FUNCTION_BLOCK FB_CIP_Source EXTENDS FB_SFC_Cycle IMPLEMENTS ITF_FB_SFC_Cycle
VAR_INPUT
	//eElementID			: E_Element_List;
	
	valTank_Water			: E_Pis_Name;
	valTank_R_Water			: E_Pis_Name;
	valTank_Detergent		: E_Pis_Name;
	valTank_DisInfection	: E_Pis_Name;	
	valDrain				: E_Pis_Name;
END_VAR
VAR_OUTPUT
END_VAR
VAR
	//refElement		: REFERENCE TO FB_Element;
	//refState_Long		: REFERENCE TO E_Element_State_Long;
	eReq				: E_CIP_Source;
	eProcess			: E_CIP_Source;
	eStatus				: E_CIP_Source;
	
	fbPis					: FB_Piston;
	stPis_Tank_Water		: REFERENCE TO ST_Piston;
	stPis_Tank_R_Water		: REFERENCE TO ST_Piston;
	stPis_Tank_Detergent	: REFERENCE TO ST_Piston;
	stPis_Tank_DisInfection	: REFERENCE TO ST_Piston;
	stPis_Drain				: REFERENCE TO ST_Piston;
	rt_Req_Reset: R_TRIG;
END_VAR
VAR_IN_OUT


END_VAR

act_GetReference();

act_Oper();
IF NOT Init.x THEN;
	act_Status();
END_IF

m_Request_Reset(memo:=rt_Req_Reset);//

ACTION _aClose_active:
bStepDone:=FALSE;
IF TRUE 
AND eStatus=E_CIP_Source.eClose
THEN;
	bStepDone:=TRUE;
END_IF
END_ACTION

ACTION _aClose_entry:
fbPis.m_SetByRecipe(stPis:=stPis_Tank_Water, 			req:=E_Piston_Recipe_State.Release);
fbPis.m_SetByRecipe(stPis:=stPis_Tank_R_Water, 			req:=E_Piston_Recipe_State.Release);
fbPis.m_SetByRecipe(stPis:=stPis_Tank_Detergent, 		req:=E_Piston_Recipe_State.Release);
fbPis.m_SetByRecipe(stPis:=stPis_Tank_DisInfection, 	req:=E_Piston_Recipe_State.Release);
fbPis.m_SetByRecipe(stPis:=stPis_Drain, 				req:=E_Piston_Recipe_State.Release);
END_ACTION

ACTION _aDetergent_entry:
fbPis.m_SetByRecipe(stPis:=stPis_Tank_Water, 			req:=E_Piston_Recipe_State.Release);
fbPis.m_SetByRecipe(stPis:=stPis_Tank_R_Water, 			req:=E_Piston_Recipe_State.Release);
fbPis.m_SetByRecipe(stPis:=stPis_Tank_Detergent, 		req:=E_Piston_Recipe_State.Act);
fbPis.m_SetByRecipe(stPis:=stPis_Tank_DisInfection, 	req:=E_Piston_Recipe_State.Release);
//fbPis.m_SetByRecipe(stPis:=stPis_Drain, 				req:=E_Piston_Recipe_State.Act);
END_ACTION

ACTION _aDone_entry:
eProcess:=E_CIP_Source.eNone;
eReq:=E_CIP_Source.eNone;
bRun:=FALSE;
bDone:=TRUE;
END_ACTION

ACTION _aInit_active:
SFCReset:=FALSE;
END_ACTION

ACTION _aInit_exit:
eProcess:=E_CIP_Source.eNone;
eReq:=E_CIP_Source.eNone;
END_ACTION

ACTION _aR_Water_entry:
fbPis.m_SetByRecipe(stPis:=stPis_Tank_Water, 			req:=E_Piston_Recipe_State.Release);
fbPis.m_SetByRecipe(stPis:=stPis_Tank_R_Water, 			req:=E_Piston_Recipe_State.Act);
fbPis.m_SetByRecipe(stPis:=stPis_Tank_Detergent, 		req:=E_Piston_Recipe_State.Release);
fbPis.m_SetByRecipe(stPis:=stPis_Tank_DisInfection, 	req:=E_Piston_Recipe_State.Release);
//fbPis.m_SetByRecipe(stPis:=stPis_Drain, 				req:=E_Piston_Recipe_State.Act);
END_ACTION

ACTION _aReady_active:


CASE eReq OF
	E_CIP_Source.eClose:;
			IF TRUE THEN;
				eProcess:=E_CIP_Source.eClose;
			END_IF

	E_CIP_Source.eT91_Sanitation:;
			IF TRUE THEN;
				eProcess:=E_CIP_Source.eT91_Sanitation;
			END_IF	
			
	E_CIP_Source.eT92_Detergent:;
			IF TRUE THEN;
				eProcess:=E_CIP_Source.eT92_Detergent;
			END_IF	

	E_CIP_Source.eT93_R_Water:;
			IF TRUE THEN;
				eProcess:=E_CIP_Source.eT93_R_Water;
			END_IF	
			
	E_CIP_Source.eT94_Water:;
			IF TRUE THEN;
				eProcess:=E_CIP_Source.eT94_Water;
			END_IF	

END_CASE
END_ACTION

ACTION _aReady_entry:

END_ACTION

ACTION _aReady_exit:
bRun:=TRUE;
bDone:=FALSE;
END_ACTION

ACTION _aSanitation_entry:
fbPis.m_SetByRecipe(stPis:=stPis_Tank_Water, 			req:=E_Piston_Recipe_State.Release);
fbPis.m_SetByRecipe(stPis:=stPis_Tank_R_Water, 			req:=E_Piston_Recipe_State.Release);
fbPis.m_SetByRecipe(stPis:=stPis_Tank_Detergent, 		req:=E_Piston_Recipe_State.Release);
fbPis.m_SetByRecipe(stPis:=stPis_Tank_DisInfection, 	req:=E_Piston_Recipe_State.Act);
END_ACTION

ACTION _aT91_Drain_Done_active:
bStepDone:=FALSE;
IF TRUE 
AND eStatus=E_CIP_Source.eT91_Sanitation
THEN;
	bStepDone:=TRUE;
END_IF
END_ACTION

ACTION _aT91_Drain_Done_entry:
fbPis.m_SetByRecipe(stPis:=stPis_Drain, 				req:=E_Piston_Recipe_State.Act);
END_ACTION

ACTION _aT92_Drain_Done_active:
bStepDone:=FALSE;
IF TRUE 
AND eStatus=E_CIP_Source.eT92_Detergent
THEN;
	bStepDone:=TRUE;
END_IF
END_ACTION

ACTION _aT92_Drain_Done_entry:
fbPis.m_SetByRecipe(stPis:=stPis_Drain, 				req:=E_Piston_Recipe_State.Act);
END_ACTION

ACTION _aT93_Drain_Done_active:
bStepDone:=FALSE;
IF TRUE 
AND eStatus=E_CIP_Source.eT93_R_Water
THEN;
	bStepDone:=TRUE;
END_IF
END_ACTION

ACTION _aT93_Drain_Done_entry:
fbPis.m_SetByRecipe(stPis:=stPis_Drain, 				req:=E_Piston_Recipe_State.Act);
END_ACTION

ACTION _aWater_active:
bStepDone:=FALSE;
IF TRUE 
AND eStatus=E_CIP_Source.eT94_Water
THEN;
	bStepDone:=TRUE;
END_IF
END_ACTION

ACTION _aWater_entry:
fbPis.m_SetByRecipe(stPis:=stPis_Tank_Water, 			req:=E_Piston_Recipe_State.Act);
fbPis.m_SetByRecipe(stPis:=stPis_Tank_R_Water, 			req:=E_Piston_Recipe_State.Release);
fbPis.m_SetByRecipe(stPis:=stPis_Tank_Detergent, 		req:=E_Piston_Recipe_State.Release);
fbPis.m_SetByRecipe(stPis:=stPis_Tank_DisInfection, 	req:=E_Piston_Recipe_State.Release);
fbPis.m_SetByRecipe(stPis:=stPis_Drain, 				req:=E_Piston_Recipe_State.Release);
END_ACTION

ACTION act_GetReference:
m_Set_SFCFlags_Reference();
//refElement REF= fbElement[eElementID];
//refState_Long REF= fbElement[eElementID].eState_Long;
	
stPis_Tank_Water			REF= g_Piston.stPis[valTank_Water];
stPis_Tank_R_Water			REF= g_Piston.stPis[valTank_R_Water];
stPis_Tank_Detergent		REF= g_Piston.stPis[valTank_Detergent];
stPis_Tank_DisInfection		REF= g_Piston.stPis[valTank_DisInfection];
stPis_Drain					REF= g_Piston.stPis[valDrain];
END_ACTION

ACTION act_Oper:
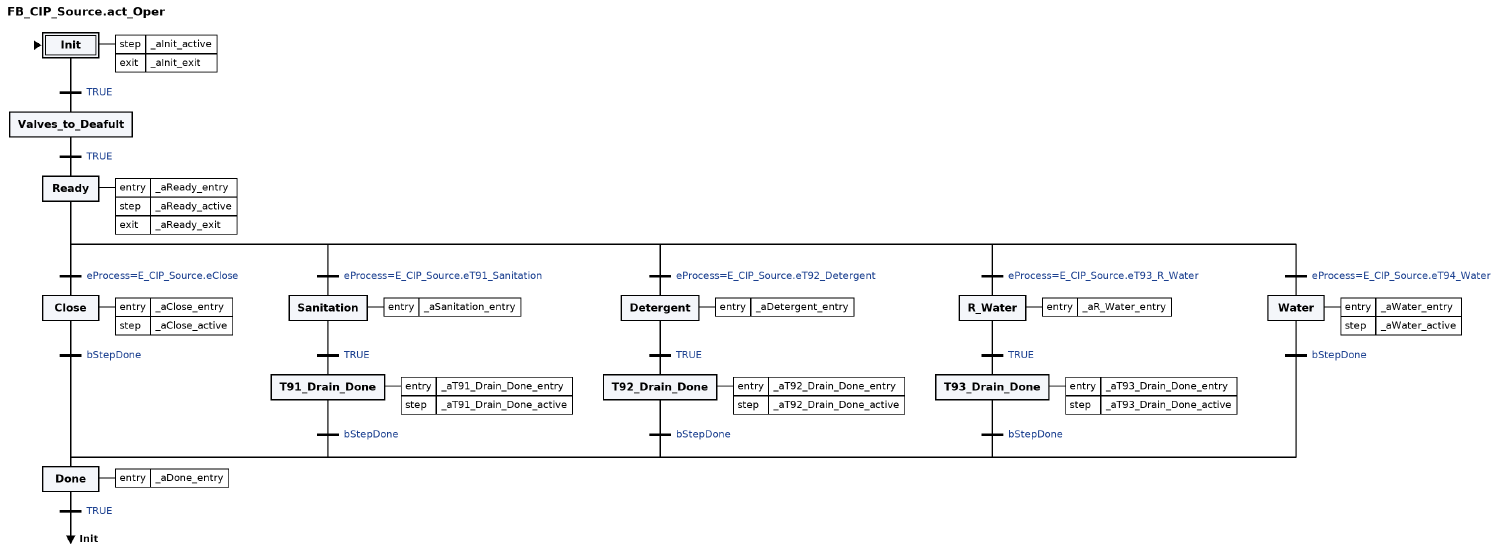
INITIAL_STEP Init:  // min time T#0.5s
    _aInit_active(N);  // step action
    _aInit_exit(P0);  // exit action
END_STEP
TRANSITION FROM Init TO Valves_to_Deafult
    := TRUE;
END_TRANSITION
STEP Valves_to_Deafult:
END_STEP
TRANSITION FROM Valves_to_Deafult TO Ready
    := TRUE;
END_TRANSITION
STEP Ready:
    _aReady_entry(P1);  // entry action
    _aReady_active(N);  // step action
    _aReady_exit(P0);  // exit action
END_STEP
TRANSITION FROM Ready TO Close
    := eProcess=E_CIP_Source.eClose;
END_TRANSITION
STEP Close:
    _aClose_entry(P1);  // entry action
    _aClose_active(N);  // step action
END_STEP
TRANSITION FROM Close TO Done
    := bStepDone;
END_TRANSITION
TRANSITION FROM Ready TO Sanitation
    := eProcess=E_CIP_Source.eT91_Sanitation;
END_TRANSITION
STEP Sanitation:  // min time T#7s
    _aSanitation_entry(P1);  // entry action
END_STEP
TRANSITION FROM Sanitation TO T91_Drain_Done
    := TRUE;
END_TRANSITION
STEP T91_Drain_Done:
    _aT91_Drain_Done_entry(P1);  // entry action
    _aT91_Drain_Done_active(N);  // step action
END_STEP
TRANSITION FROM T91_Drain_Done TO Done
    := bStepDone;
END_TRANSITION
TRANSITION FROM Ready TO Detergent
    := eProcess=E_CIP_Source.eT92_Detergent;
END_TRANSITION
STEP Detergent:  // min time T#6s
    _aDetergent_entry(P1);  // entry action
END_STEP
TRANSITION FROM Detergent TO T92_Drain_Done
    := TRUE;
END_TRANSITION
STEP T92_Drain_Done:
    _aT92_Drain_Done_entry(P1);  // entry action
    _aT92_Drain_Done_active(N);  // step action
END_STEP
TRANSITION FROM T92_Drain_Done TO Done
    := bStepDone;
END_TRANSITION
TRANSITION FROM Ready TO R_Water
    := eProcess=E_CIP_Source.eT93_R_Water;
END_TRANSITION
STEP R_Water:  // min time T#5s
    _aR_Water_entry(P1);  // entry action
END_STEP
TRANSITION FROM R_Water TO T93_Drain_Done
    := TRUE;
END_TRANSITION
STEP T93_Drain_Done:
    _aT93_Drain_Done_entry(P1);  // entry action
    _aT93_Drain_Done_active(N);  // step action
END_STEP
TRANSITION FROM T93_Drain_Done TO Done
    := bStepDone;
END_TRANSITION
TRANSITION FROM Ready TO Water
    := eProcess=E_CIP_Source.eT94_Water;
END_TRANSITION
STEP Water:
    _aWater_entry(P1);  // entry action
    _aWater_active(N);  // step action
END_STEP
TRANSITION FROM Water TO Done
    := bStepDone;
END_TRANSITION
STEP Done:  // min time T#0.2s
    _aDone_entry(P1);  // entry action
END_STEP
TRANSITION FROM Done TO Init
    := TRUE;
END_TRANSITION
// branch label Branch1_act_Oper
END_ACTION

ACTION act_Status:
IF bReady AND bDone OR TRUE THEN;
	IF TRUE 
	AND fbPis.m_CheckByRecipe(stPis:=stPis_Tank_Water, 			req:=E_Piston_Recipe_State.Release)
	AND fbPis.m_CheckByRecipe(stPis:=stPis_Tank_R_Water, 		req:=E_Piston_Recipe_State.Release)
	AND fbPis.m_CheckByRecipe(stPis:=stPis_Tank_Detergent, 		req:=E_Piston_Recipe_State.Release)
	AND fbPis.m_CheckByRecipe(stPis:=stPis_Tank_DisInfection, 	req:=E_Piston_Recipe_State.Release)
	AND fbPis.m_CheckByRecipe(stPis:=stPis_Drain, 				req:=E_Piston_Recipe_State.Release)
	THEN;
		eStatus:=E_CIP_Source.eClose;
	
	ELSIF TRUE 
	AND fbPis.m_CheckByRecipe(stPis:=stPis_Tank_Water, 			req:=E_Piston_Recipe_State.Act)
	AND fbPis.m_CheckByRecipe(stPis:=stPis_Tank_R_Water, 		req:=E_Piston_Recipe_State.Release)
	AND fbPis.m_CheckByRecipe(stPis:=stPis_Tank_Detergent, 		req:=E_Piston_Recipe_State.Release)
	AND fbPis.m_CheckByRecipe(stPis:=stPis_Tank_DisInfection, 	req:=E_Piston_Recipe_State.Release)
	AND fbPis.m_CheckByRecipe(stPis:=stPis_Drain, 				req:=E_Piston_Recipe_State.Release)
	THEN;
		eStatus:=E_CIP_Source.eT94_Water;
		
	ELSIF TRUE 
	AND fbPis.m_CheckByRecipe(stPis:=stPis_Tank_Water, 			req:=E_Piston_Recipe_State.Release)
	AND fbPis.m_CheckByRecipe(stPis:=stPis_Tank_R_Water, 		req:=E_Piston_Recipe_State.Act)
	AND fbPis.m_CheckByRecipe(stPis:=stPis_Tank_Detergent, 		req:=E_Piston_Recipe_State.Release)
	AND fbPis.m_CheckByRecipe(stPis:=stPis_Tank_DisInfection, 	req:=E_Piston_Recipe_State.Release)
	AND fbPis.m_CheckByRecipe(stPis:=stPis_Drain, 				req:=E_Piston_Recipe_State.Act)
	THEN;
		eStatus:=E_CIP_Source.eT93_R_Water;
		
	ELSIF TRUE 	
	AND fbPis.m_CheckByRecipe(stPis:=stPis_Tank_Water, 			req:=E_Piston_Recipe_State.Release)
	AND fbPis.m_CheckByRecipe(stPis:=stPis_Tank_R_Water, 		req:=E_Piston_Recipe_State.Release)
	AND fbPis.m_CheckByRecipe(stPis:=stPis_Tank_Detergent, 		req:=E_Piston_Recipe_State.Act)
	AND fbPis.m_CheckByRecipe(stPis:=stPis_Tank_DisInfection, 	req:=E_Piston_Recipe_State.Release)
	AND fbPis.m_CheckByRecipe(stPis:=stPis_Drain, 				req:=E_Piston_Recipe_State.Act)
	THEN;
		eStatus:=E_CIP_Source.eT92_Detergent;
		
	ELSIF TRUE 	
	AND fbPis.m_CheckByRecipe(stPis:=stPis_Tank_Water, 			req:=E_Piston_Recipe_State.Release)
	AND fbPis.m_CheckByRecipe(stPis:=stPis_Tank_R_Water, 		req:=E_Piston_Recipe_State.Release)
	AND fbPis.m_CheckByRecipe(stPis:=stPis_Tank_Detergent, 		req:=E_Piston_Recipe_State.Release)
	AND fbPis.m_CheckByRecipe(stPis:=stPis_Tank_DisInfection, 	req:=E_Piston_Recipe_State.Act)
	AND fbPis.m_CheckByRecipe(stPis:=stPis_Drain, 				req:=E_Piston_Recipe_State.Act)
	THEN;
		eStatus:=E_CIP_Source.eT91_Sanitation;
	ELSE;
		eStatus:=E_Tank_Target.eNone;
	END_IF
ELSE;
	eStatus:=E_Tank_Target.eNone;
END_IF
END_ACTION

METHOD m_CheckStatus : BOOL
VAR_INPUT
	eReqStatus		: E_CIP_Source;
END_VAR
IF eStatus=eReqStatus 
AND eProcess=E_CIP_Source.eNone
AND eReq=E_CIP_Source.eNone
AND bReady
AND bDone
AND NOT bRun
THEN;
	m_CheckStatus:=TRUE;
END_IF
END_METHOD

METHOD m_Request_Reset : BOOL
VAR_IN_OUT
	memo: R_TRIG;
END_VAR
memo(CLK:=eReq=0);
IF TRUE 
AND memo.Q
THEN;
	SFCReset:=TRUE;
END_IF
END_METHOD

METHOD m_Run : BOOL
VAR_INPUT
	eReqProc			: E_CIP_Source;
END_VAR
IF eProcess=E_CIP_Source.eNone THEN;
	eProcess:=eReq:=eReqProc;
	bDone:=FALSE;
	m_Run:=TRUE;
END_IF
END_METHOD

METHOD m_Set_SFCFlags_Reference : BOOL
//Set reference to SFC flags

refSFC.SFCInit REF= SFCInit;
refSFC.SFCReset REF= SFCReset;
refSFC.SFCError REF= SFCError;
refSFC.SFCEnableLimit REF= SFCEnableLimit;
refSFC.SFCErrorStep REF= SFCErrorStep;
refSFC.SFCErrorPOU REF= SFCErrorPOU;
refSFC.SFCQuitError REF= SFCQuitError;
refSFC.SFCPause REF= SFCPause;
refSFC.SFCTrans REF= SFCTrans;
refSFC.SFCCurrentStep REF= SFCCurrentStep;
refSFC.SFCTip REF= SFCTip;
refSFC.SFCTipMode REF= SFCTipMode;

// Cycle handle for SFC
m_SFC_Handle();
END_METHOD

END_FUNCTION_BLOCK

(* stored: Version 1.1.0.1, ProductVersion 3.1.4024.13
   POU FB_CIP_Source: Id {51aff4c3-d299-4189-9ddb-b537da8ea506}, SpecialFunc None
   Folder Manage: Id {f72c9a77-5990-4e2a-906f-d727cb28c56e}
   Action _aClose_active: Id {31213e26-c963-4ed4-8ec0-5daeea10e078}
   Action _aClose_entry: Id {d09c7332-d193-4493-b1e4-5232db477b55}
   Action _aDetergent_entry: Id {771716ff-47a9-481a-a6f9-85f73c1e2b6e}
   Action _aDone_entry: Id {d6158c19-8f25-4535-8bf6-7e51dd1b5362}
   Action _aInit_active: Id {1f5ddc3a-233c-4a03-b1ef-5e34b8a9ca83}
   Action _aInit_exit: Id {f16fd208-cc2f-42cd-a16b-26e036360a07}
   Action _aR_Water_entry: Id {4de374b9-bbb5-4b70-9cc6-a1672e94772e}
   Action _aReady_active: Id {2f0857dc-1162-4f85-849b-826c1f096529}
   Action _aReady_entry: Id {504413b8-8cea-4dae-9c16-ea892c8ff1ad}
   Action _aReady_exit: Id {4a59497c-bd7d-4bd0-bb0d-43d900603e02}
   Action _aSanitation_entry: Id {3930e00c-3e06-4f7e-94da-486d833daa71}
   Action _aT91_Drain_Done_active: Id {f4899e9e-1998-4384-be9f-6b66921960ee}
   Action _aT91_Drain_Done_entry: Id {54a143b9-5f4f-4124-8530-071d5d31260e}
   Action _aT92_Drain_Done_active: Id {e74836d7-8079-4924-8aa7-ad2028b472cc}
   Action _aT92_Drain_Done_entry: Id {0ba5c126-6f68-4257-b981-8742b6a006cb}
   Action _aT93_Drain_Done_active: Id {a28d0589-c36e-4ff5-a15c-aa7370ba98c4}
   Action _aT93_Drain_Done_entry: Id {8dbcb274-8858-4ef1-a4ef-1408fe354ee9}
   Action _aWater_active: Id {b975f465-2f2b-45f4-b094-9a9c16edef44}
   Action _aWater_entry: Id {597c2d38-8971-4aaa-9c62-38b287ee2e35}
   Action act_GetReference: Id {553e7d71-99a7-47aa-ae6f-0cd5ac38902f}
   Action act_Oper: Id {5af8f4ab-bced-408d-828d-06e969601154}
   Action act_Status: Id {8c5bd8f8-66f0-4098-9f33-9015434f732a}
   Method m_CheckStatus: Id {cc574672-75d4-4109-af68-d1c872851152}
   Method m_Request_Reset: Id {54a4460d-5097-43de-b69e-b82abb168d84}
   Method m_Run: Id {5d191ab6-be10-46af-8016-5701543b152c}
   Method m_Set_SFCFlags_Reference: Id {6a5e32bd-46a1-4d83-b2b2-41e90d72387a} *)
